(* PLC project Vn_member_assign, Beckhoff Automation GmbH TwinCAT PLC Control 3.5.13.21 *)
(* stored: creationDateTime 1970-01-01T00:00:00 *)

PROGRAM Vn_member_assign

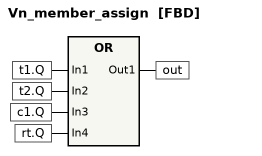
(* FBD diagram, written out as Structured Text *)
out := t1.Q OR t2.Q OR c1.Q OR rt.Q;
END_PROGRAM
